(* CODESYS project id.library
   DefaultNamespace: KOSTAL.AF2024.Core.ID
   DocFormat: reStructuredText
   Description: Base Library for identifier functions (Index + Name)
   Author: Frank Dümpelmann
   Title: KOSTAL.AF2024.Core.ID
   Version: 1.0.0.0
   Company: KOSTAL GmbH & Co.KG
   Placeholder: KOSTAL.AF2024.Core.ID

Project tree, tasks and I/O mapping:
  libraries: KOSTAL.AF2024.Core.Settings, 1.0.0.0 (KOSTAL GmbH & Co.KG); KOSTAL.AF2024.Core.System, 1.0.0.0 (KOSTAL GmbH & Co.KG)
  DUT/
    interface I_T_ID: CopyTo, key, name
    interface I_T_ID_CopyFrom: CopyFrom
    interface I_T_ID_Owner: clear, CopyFrom, CopyTo, key, name
    function block T_ID [ST]: clear, CopyFrom, CopyTo, key, name
  Project Information/
    function F_GetCompany [ST]
    function F_GetTitle [ST]
    function F_GetVersion [ST]
  Version/
    global variables Global_Version
*)

// Version/Global_Version
{attribute 'TcGenerated'}
{attribute 'no-analysis'}
{attribute 'linkalways'}
// This function has been automatically generated from the project information.
VAR_GLOBAL CONSTANT
	{attribute 'const_non_replaced'}
	stLibVersion_KOSTAL_AF2024_Core_ID : ST_LibVersion := (iMajor := 1, iMinor := 0, iBuild := 0, iRevision := 0, nFlags := 0, sVersion := '1.0.0.0');
END_VAR

// DUT/I_T_ID
INTERFACE I_T_ID EXTENDS KOSTAL_AF2024_Core_System.I_Interface

METHOD PUBLIC CopyTo
VAR_INPUT
	IN	:	I_T_ID_CopyFrom;
END_VAR
END_METHOD

PROPERTY PUBLIC key : DINT
GET
END_GET
END_PROPERTY

PROPERTY PUBLIC name : KOSTAL_AF2024_Core_Settings.T_MaxString
GET
END_GET
END_PROPERTY

END_INTERFACE

// DUT/I_T_ID_CopyFrom
INTERFACE I_T_ID_CopyFrom EXTENDS KOSTAL_AF2024_Core_System.I_Interface

METHOD PUBLIC CopyFrom
VAR_INPUT
	IN	: I_T_ID;
END_VAR
END_METHOD

END_INTERFACE

// DUT/I_T_ID_Owner
INTERFACE I_T_ID_Owner EXTENDS KOSTAL_AF2024_Core_System.I_Interface

METHOD PUBLIC clear
VAR_INPUT
END_VAR
END_METHOD

METHOD PUBLIC CopyFrom
VAR_INPUT
	IN	: I_T_ID;
END_VAR
END_METHOD

METHOD PUBLIC CopyTo
VAR_INPUT
	IN	:	I_T_ID_CopyFrom;
END_VAR
END_METHOD

PROPERTY PUBLIC key : DINT
GET
END_GET
SET
END_SET
END_PROPERTY

PROPERTY PUBLIC name : KOSTAL_AF2024_Core_Settings.T_MaxString
GET
END_GET
SET
END_SET
END_PROPERTY

END_INTERFACE

// DUT/T_ID
(*

:Author: Frank Dümpelmann <f.duempelmann@kostal.com>
:Date: 2018-10-19

Function
========
Base data structure for identifier functions (Index + Name)

*)
{attribute 'enable_dynamic_creation'}
FUNCTION_BLOCK PUBLIC T_ID IMPLEMENTS I_T_ID, I_T_ID_CopyFrom, I_T_ID_Owner

VAR
		_key 	: DINT;
		_name	: KOSTAL_AF2024_Core_Settings.T_MaxString;
END_VAR

METHOD PUBLIC clear
VAR_INPUT
END_VAR

_key	:= 0;
_name	:= "";
END_METHOD

METHOD PUBLIC CopyFrom
VAR_INPUT
	IN	: I_T_ID;
END_VAR

IF IN = 0 THEN	RETURN;	END_IF

_key	:= IN.key;
_name	:= IN.name;
END_METHOD

METHOD PUBLIC CopyTo
VAR_INPUT
	IN	:	I_T_ID_CopyFrom;
END_VAR

IF IN = 0 THEN	RETURN;	END_IF

IN.CopyFrom(THIS^);
END_METHOD

PROPERTY PUBLIC key : DINT
GET

key:= _key;
END_GET
SET

_key:= key;
END_SET
END_PROPERTY

PROPERTY PUBLIC name : KOSTAL_AF2024_Core_Settings.T_MaxString
GET

name := _name;
END_GET
SET

_name := name;
END_SET
END_PROPERTY

END_FUNCTION_BLOCK

// Project Information/F_GetCompany
// This function has been automatically generated from the project information.
{attribute 'signature_flag' := '1073741824'}
{attribute 'TcGenerated'}
{attribute 'no-analysis'}
FUNCTION F_GetCompany : WSTRING
VAR_INPUT
	
END_VAR

F_GetCompany := "KOSTAL GmbH & Co.KG";

END_FUNCTION

// Project Information/F_GetTitle
// This function has been automatically generated from the project information.
{attribute 'signature_flag' := '1073741824'}
{attribute 'TcGenerated'}
{attribute 'no-analysis'}
FUNCTION F_GetTitle : WSTRING
VAR_INPUT
	
END_VAR

F_GetTitle := "KOSTAL.AF2024.Core.ID";

END_FUNCTION

// Project Information/F_GetVersion
// This function has been automatically generated from the project information.
{attribute 'signature_flag' := '1073741824'}
{attribute 'TcGenerated'}
{attribute 'no-analysis'}
FUNCTION F_GetVersion : ST_LibVersion
VAR_INPUT
	
END_VAR

F_GetVersion.iMajor := 1;
F_GetVersion.iMinor := 0;
F_GetVersion.iBuild := 0;
F_GetVersion.iRevision := 0;
F_GetVersion.sVersion := '1.0.0.0';
F_GetVersion.nFlags := 0;

END_FUNCTION
